Fanuc KAREL source: KB00156.KL

PROGRAM KB00156
%NOLOCKGROUP
%ENVIRONMENT TPE
VAR
  P1: STRING[80]
  P2: INTEGER
BEGIN
  P1 = 'A'
  P2 = 1
  SELECT_TPE(P1, P2)
END KB00156
